Fanuc KAREL source: KC00009.KL

PROGRAM KC00009
%NOLOCKGROUP
%ENVIRONMENT PATHOP
VAR
  I: INTEGER
  J: INTEGER
  K: INTEGER
  R: REAL
  B: BOOLEAN
  S: STRING[80]
  T: STRING[80]
  P: PATH
  Q: PATH
  AI: ARRAY[8] OF INTEGER
  AB: ARRAY[244] OF BYTE
BEGIN
  INSERT_NODE(P,I,J)
END KC00009
